KUKA KRL data list: folge11.dat

&ACCESS RVP
&REL 1
&COMMENT bt2krl vw-ks24 data Folge 11 plan 16#A1BE
DEFDAT FOLGE11
   ; Generated by bt2krl 0.1.0 from bt2plc plan bt_1792156523_scene_fit (cell scene_fit), PLAN_ID 16#A1BE
   ; Robot robot1 (R1), controller robot1, model unknown, joint mapping identity
   ; Profile vw-ks24 (VW KS24 / TPVW 8.1.8).
   ; Do not edit: regenerate with bt2krl (plain KRL, no inline forms).
   EXT BAS (BAS_COMMAND :IN,REAL :IN )
   ; interface to the VW standard routines (as every VW Folge .dat declares them)
   EXT VW (VW_COMMAND :IN,BOOL :IN,REAL :IN,REAL :IN,REAL :IN,REAL :IN,BOOL :IN,E6POS :IN )
   EXT VW_USR_R (VW_USER_CMD :IN,INT :IN,REAL :IN,REAL :IN,REAL :IN,REAL :IN,REAL :IN,REAL :IN,BOOL :IN )
   EXTFCT INT SELECT (SUBTYPE :IN,INT :IN,BOOL :IN,ARI_TYP :IN,INT :IN,BOOL_TYP :IN,INT :IN,BOOL :IN)
   DECL AXIS P0={A1 45.0,A2 -90.0,A3 90.0,A4 0.0,A5 0.0,A6 0.0}
   DECL AXIS P1={A1 43.6012,A2 -89.7676,A3 90.0033,A4 0.0,A5 1.8605,A6 -0.3507}
   DECL AXIS P2={A1 41.9543,A2 -89.4939,A3 90.0071,A4 0.0,A5 4.051,A6 -0.7636}
   DECL AXIS P3={A1 37.1038,A2 -88.6879,A3 90.0185,A4 0.0,A5 10.5026,A6 -1.9796}
   DECL AXIS P4={A1 26.9514,A2 -87.001,A3 90.0423,A4 0.0,A5 24.006,A6 -4.5249}
   DECL AXIS P5={A1 6.8724,A2 -83.6646,A3 90.0893,A4 0.0,A5 50.7127,A6 -9.5588}
   DECL AXIS P6={A1 -4.0921,A2 -81.8426,A3 90.115,A4 0.0,A5 65.2964,A6 -12.3077}
   DECL AXIS P7={A1 -9.8225,A2 -80.8905,A3 90.1284,A4 0.0,A5 72.9183,A6 -13.7444}
   DECL AXIS P8={A1 -12.0109,A2 -80.5268,A3 90.1336,A4 0.0,A5 75.829,A6 -14.293}
   DECL AXIS P9={A1 -14.6956,A2 -80.0807,A3 90.1398,A4 0.0,A5 79.3999,A6 -14.9661}
   DECL AXIS P10={A1 -15.0566,A2 -80.0207,A3 90.1407,A4 0.0,A5 79.88,A6 -15.0566}
   DECL AXIS P11={A1 -15.0566,A2 -79.875,A3 90.7142,A4 0.0,A5 79.1607,A6 -15.0566}
   DECL AXIS P12={A1 -15.0566,A2 -79.6592,A3 91.5498,A4 0.0,A5 78.1094,A6 -15.0566}
   DECL AXIS P13={A1 -15.0566,A2 -78.7933,A3 94.228,A4 0.0,A5 74.5653,A6 -15.0566}
   DECL AXIS P14={A1 -15.0374,A2 -79.913,A3 90.5893,A4 0.0,A5 79.3237,A6 -15.0374}
   DECL AXIS P15={A1 -13.7654,A2 -80.0274,A3 90.142,A4 0.0,A5 79.8854,A6 -13.7654}
   DECL AXIS P16={A1 -9.2939,A2 -80.052,A3 90.1253,A4 0.0,A5 79.9267,A6 -9.2939}
   DECL AXIS P17={A1 8.1168,A2 -80.1118,A3 90.221,A4 0.0,A5 79.8908,A6 8.1168}
   DECL AXIS P18={A1 11.5499,A2 -80.1218,A3 90.2471,A4 0.0,A5 79.8747,A6 11.5498}
   DECL AXIS P19={A1 13.8795,A2 -80.1284,A3 90.2658,A4 0.0,A5 79.8625,A6 13.8794}
   DECL AXIS P20={A1 14.7377,A2 -80.1307,A3 90.273,A4 0.0,A5 79.8577,A6 14.7377}
   DECL AXIS P21={A1 14.7377,A2 -79.9847,A3 90.8466,A4 0.0,A5 79.1381,A6 14.7377}
   DECL AXIS P22={A1 14.7377,A2 -79.7685,A3 91.6823,A4 0.0,A5 78.0862,A6 14.7377}
   DECL AXIS P23={A1 14.7377,A2 -78.9012,A3 94.361,A4 0.0,A5 74.5402,A6 14.7377}
   DECL AXIS P24={A1 14.7377,A2 -79.9556,A3 90.9835,A4 0.0,A5 78.9721,A6 14.7377}
   DECL AXIS P25={A1 15.0076,A2 -80.0451,A3 90.9747,A4 0.0,A5 78.2679,A6 14.6063}
   DECL AXIS P26={A1 15.7755,A2 -80.3,A3 90.9498,A4 0.0,A5 76.2638,A6 14.2323}
   DECL AXIS P27={A1 16.9794,A2 -80.6996,A3 90.9106,A4 0.0,A5 73.1223,A6 13.646}
   DECL AXIS P28={A1 18.5568,A2 -81.2232,A3 90.8594,A4 0.0,A5 69.0058,A6 12.8778}
   DECL AXIS P29={A1 22.5835,A2 -82.5597,A3 90.7285,A4 0.0,A5 58.4978,A6 10.9168}
   DECL AXIS P30={A1 34.8296,A2 -86.6243,A3 90.3305,A4 0.0,A5 26.5407,A6 4.953}
   DECL AXIS P31={A1 39.2921,A2 -88.1055,A3 90.1855,A4 0.0,A5 14.8953,A6 2.7797}
   DECL AXIS P32={A1 41.1809,A2 -88.7324,A3 90.1241,A4 0.0,A5 9.9663,A6 1.8599}
   DECL AXIS P33={A1 43.9622,A2 -89.6555,A3 90.0337,A4 0.0,A5 2.7082,A6 0.5054}
   DECL AXIS P34={A1 44.7302,A2 -89.9104,A3 90.0088,A4 0.0,A5 0.7041,A6 0.1314}
   DECL AXIS P35={A1 45.0,A2 -90.0,A3 90.0,A4 0.0,A5 0.0,A6 0.0}
ENDDAT
